FUNCTION_BLOCK FB_Error_Handle
VAR_INPUT
	bError: BOOL;
	sErrID: STRING;
END_VAR
VAR_OUTPUT
END_VAR
VAR
	fbFormat: FB_FormatString;
END_VAR
VAR_IN_OUT
	error_code: STRING;

END_VAR



IF bError 
AND error_code=''
THEN;
	error_code:=sErrID;
END_IF

IF NOT bError 
AND error_code=sErrID
THEN;
	error_code:='';
END_IF

METHOD m_GetAxisErr : STRING(4)
VAR_INPUT
	stDevErr_H				: ST_DeviceErrorHandeling;
END_VAR
VAR_OUTPUT
	sMessage: STRING;
END_VAR

VAR
	ErrID_xx: STRING(2);
END_VAR
IF bError 
AND error_code=''
THEN;
	fbFormat(sFormat:='%0.2d' ,arg1:=F_INT(stDevErr_H.iObjectID),sOut=>ErrID_xx);
	m_GetAxisErr:=CONCAT('23',ErrID_xx);
	sMessage:=stDevErr_H.sObjectName;
ELSE;
	m_GetAxisErr:='';
END_IF
END_METHOD

METHOD m_GetPistonErr : STRING(4)
VAR_INPUT
	stDevErr_H				: ST_DeviceErrorHandeling;
END_VAR
VAR_OUTPUT
	sMessage: STRING;
END_VAR

VAR
	ErrID_xx: STRING(2);
END_VAR
IF bError 
AND error_code=''
THEN;
	fbFormat(sFormat:='%0.2d' ,arg1:=F_INT(stDevErr_H.iObjectID),sOut=>ErrID_xx);
	m_GetPistonErr:=CONCAT('22',ErrID_xx);
	sMessage:=stDevErr_H.sObjectName;
ELSE;
	m_GetPistonErr:='';
END_IF
END_METHOD

END_FUNCTION_BLOCK

(* stored: Version 1.1.0.1, ProductVersion 3.1.4024.12
   POU FB_Error_Handle: Id {b9c0feb5-6ac8-4d06-98ea-e57922381035}, SpecialFunc None
   Method m_GetAxisErr: Id {fdcaa3bf-1b97-4a77-92a2-67637e90edf8}
   Method m_GetPistonErr: Id {b3c5c7fd-4af7-4524-a42c-4563611997f1} *)
